(* IEC 61131-3 sources: plc-st-coding-agent/progress/f14_agent_v4_diagnostics/release/review/f14_self, 2 files *)

(* ---- fill_codex_deepseek-v4pro.st ---- *)
FUNCTION_BLOCK FB
VAR_INPUT
    startBtn : BOOL;
    resetBtn : BOOL;
    doneSensor : BOOL;
    targetVol : REAL;
    flowVol : REAL;
END_VAR
VAR_OUTPUT
    valveOpen : BOOL;
    fillsToday : INT;
END_VAR
VAR
    accVol : REAL;
    pendingConfirm : BOOL;
    startPrev : BOOL;
    resetPrev : BOOL;
    startRising : BOOL;
    resetRising : BOOL;
    valveWasOpen : BOOL;
END_VAR

startRising := startBtn AND NOT startPrev;
resetRising := resetBtn AND NOT resetPrev;
valveWasOpen := valveOpen;

IF resetRising THEN
    valveOpen := FALSE;
    fillsToday := 0;
    accVol := 0.0;
    pendingConfirm := FALSE;

ELSIF startRising AND NOT valveWasOpen THEN
    accVol := flowVol;
    valveOpen := accVol < targetVol;
    pendingConfirm := NOT valveOpen;

ELSIF valveWasOpen THEN
    accVol := accVol + flowVol;
    IF accVol < targetVol THEN
        valveOpen := TRUE;
        pendingConfirm := FALSE;
    ELSE
        valveOpen := FALSE;
        pendingConfirm := TRUE;
    END_IF

ELSIF pendingConfirm THEN
    valveOpen := FALSE;
    IF doneSensor THEN
        IF fillsToday < 32767 THEN
            fillsToday := fillsToday + 1;
        END_IF
        pendingConfirm := FALSE;
        accVol := 0.0;
    END_IF

ELSE
    valveOpen := FALSE;
    pendingConfirm := FALSE;
    accVol := 0.0;
END_IF

startPrev := startBtn;
resetPrev := resetBtn;

END_FUNCTION_BLOCK

(* ---- fill_custom_deepseek-v4pro.st ---- *)
FUNCTION_BLOCK FB
VAR_INPUT
    startBtn : BOOL;
    resetBtn : BOOL;
    doneSensor : BOOL;
    targetVol : REAL;
    flowVol : REAL;
END_VAR
VAR_OUTPUT
    valveOpen : BOOL;
    fillsToday : INT;
END_VAR
VAR
    startBtn_prev : BOOL;
    resetBtn_prev : BOOL;
    is_filling : BOOL;
    accumulated_volume : REAL;
    waiting_for_done : BOOL;
    start_rising : BOOL;
    reset_rising : BOOL;
END_VAR

start_rising := startBtn AND NOT startBtn_prev;
reset_rising := resetBtn AND NOT resetBtn_prev;

IF reset_rising THEN
    fillsToday := 0;
    valveOpen := FALSE;
    accumulated_volume := 0.0;
    waiting_for_done := FALSE;
    is_filling := FALSE;
ELSE
    IF start_rising AND NOT is_filling THEN
        waiting_for_done := FALSE;
        is_filling := TRUE;
        accumulated_volume := 0.0;
    END_IF;

    IF is_filling THEN
        accumulated_volume := accumulated_volume + flowVol;
        IF accumulated_volume >= targetVol THEN
            valveOpen := FALSE;
            is_filling := FALSE;
            waiting_for_done := TRUE;
        ELSE
            valveOpen := TRUE;
        END_IF;
    ELSE
        valveOpen := FALSE;
        IF waiting_for_done AND doneSensor THEN
            IF fillsToday < 32767 THEN
                fillsToday := fillsToday + 1;
            END_IF;
            waiting_for_done := FALSE;
        END_IF;
    END_IF;
END_IF;

startBtn_prev := startBtn;
resetBtn_prev := resetBtn;

END_FUNCTION_BLOCK
